DATA_BLOCK "DB_IO"
{ S7_Optimized_Access := 'TRUE' }
VERSION : 0.1
NON_RETAIN
   VAR
      xStartPB : Bool;
      xStopPB : Bool := TRUE;
      xOverload : Bool;
   END_VAR

BEGIN

END_DATA_BLOCK
